(* IEC 61131-3 sources: labpomirs3/AsIOTime, 3 files *)

(* ---- AsIOTime.typ ---- *)
(********************************************************************
 * COPYRIGHT -- Bernecker + Rainer
 ********************************************************************
 * Library: AsIOTime
 * File: AsIOTime.typ
 * Author: B+R
 ********************************************************************
 * Data types of library AsIOTime
 ********************************************************************)

TYPE

END_TYPE

(* ---- AsIOTime.fun ---- *)
(********************************************************************
 * COPYRIGHT -- Bernecker + Rainer
 ********************************************************************
 * Library: AsIOTime
 * File: AsIOTime.fun
 * Author: B+R
 ********************************************************************
 * Functions and function blocks of library AsIOTime
 ********************************************************************)

{REDUND_OK} {REDUND_UNREPLICABLE} FUNCTION AsIOTimeStamp : DINT (* Get current SystemTime stamp in microseconds *)
END_FUNCTION

{REDUND_CONTEXT} {REDUND_UNREPLICABLE} FUNCTION AsIOTimeCyclicStart : DINT (* Get SystemTime at start of cyclic ressource *)
END_FUNCTION

(* ---- AsIOTime.var ---- *)
(********************************************************************
 * COPYRIGHT -- Bernecker + Rainer
 ********************************************************************
 * Library: AsIOTime
 * File: AsIOTime.var
 * Author: B+R
 ********************************************************************
 * Local variables of library AsIOTime
 ********************************************************************)

VAR CONSTANT

END_VAR
